Fanuc KAREL source: KT00691.KL

PROGRAM KT00691
%NOLOCKGROUP
VAR
  V1: VECTOR
  V2: VECTOR
  OUT: INTEGER
BEGIN
  V1.X = 1.0
  V2.Y = 2.0
  V1.X = 1.0
  V2.Y = 2.0
  OUT = + V1
END KT00691
